Fanuc KAREL source: KT00428.KL

PROGRAM KT00428
%NOLOCKGROUP
VAR
  P1: XYZWPREXT
  P2: XYZWPR
  OUT: BOOLEAN
BEGIN
  P1.X = 1.0
    P2.Y = 2.0
  OUT = P1 > P2
END KT00428
